Staubli VAL3: bind.pgx

public program bind()
  local num l_i
  local string l_sbtn
begin
  //lst
  userPageBind("prog","lst1","options",sList,49,"r")
  userPageBind("prog","lst1","value",sSelProg,1,"rw")
  for l_i = 0 to size(bBool)-1
    l_sbtn="btn"+toString("",l_i)
    userPageBindClick("prog",l_sbtn,bBool[l_i],true)
  endFor
  userPageBindClick("prog","btnback",bBack,true)
  userPageBind("prog","lbleditindex","innerHTML",sPageIndex,1,"r")
  userPageBind("prog","lbleditpage","innerHTML",sPageNum,1,"r")
end
